FUNCTION_BLOCK Mixing
VAR_INPUT
	diEnabled : BOOL;
	iSecImp : BOOL;
END_VAR
VAR_OUTPUT
	doEnabled : BOOL;
END_VAR
VAR_IN_OUT
	MixingPhase : TPhaseMixing;
	MixerEng : TEngine;
END_VAR
VAR
	rtSecImp : R_TRIG;          // rising edge of second impulse
END_VAR

{region "Aut/Man"}
    // switching state of phase - automatic or manual control (default state is manual)
    // if both commands come at once, manual has priority (safety)
    IF MixingPhase.Cmd.ManCtrl THEN
        MixingPhase.State.ManCtrl := TRUE;
        MixingPhase.State.AutCtrl := FALSE;
    ELSIF MixingPhase.Cmd.AutCtrl THEN
        MixingPhase.State.ManCtrl := FALSE;
        MixingPhase.State.AutCtrl := TRUE;
    END_IF;

    // initialization - if neither mode is active, use manual
    IF NOT MixingPhase.State.AutCtrl AND NOT MixingPhase.State.ManCtrl THEN
        MixingPhase.State.ManCtrl := TRUE;
    END_IF;

    // commands are always reset after processing
    MixingPhase.Cmd.ManCtrl := FALSE;
    MixingPhase.Cmd.AutCtrl := FALSE;
{endregion}

{region "ManCtrl"}
    // processing manual actions - if command is processed, it is set to FALSE even if can't be processed
    // Phase commands are start, stop, pause and resume
    // Start  - start mixing (elapsed time starts from 0)
    // Stop   - stop mixing
    // Pause  - stop mixing (elapsed time is kept)
    // Resume - start mixing (continues for the remaining time)
    IF MixingPhase.State.ManCtrl THEN
        IF MixingPhase.State.Idle AND MixingPhase.Cmd.StartMan THEN
            MixingPhase.State.Running := TRUE;
            MixingPhase.State.Idle := FALSE;
            MixingPhase.State.Paused := FALSE;
            MixingPhase.State.Done := FALSE;
            MixingPhase.ElapsedTimeSec := 0;
        ELSIF MixingPhase.Cmd.StopMan THEN
            MixingPhase.State.Running := FALSE;
            MixingPhase.State.Idle := TRUE;
            MixingPhase.State.Paused := FALSE;
        ELSIF MixingPhase.State.Running AND MixingPhase.Cmd.PauseMan THEN
            MixingPhase.State.Running := FALSE;
            MixingPhase.State.Idle := FALSE;
            MixingPhase.State.Paused := TRUE;
        ELSIF MixingPhase.State.Paused AND MixingPhase.Cmd.ResumeMan THEN
            MixingPhase.State.Running := TRUE;
            MixingPhase.State.Idle := FALSE;
            MixingPhase.State.Paused := FALSE;
            MixingPhase.State.Done := FALSE;
        END_IF;
    END_IF;

    MixingPhase.Cmd.StartMan := FALSE;
    MixingPhase.Cmd.StopMan := FALSE;
    MixingPhase.Cmd.PauseMan := FALSE;
    MixingPhase.Cmd.ResumeMan := FALSE;
{endregion}

{region "AutCtrl"}
    // if phase is in automatic mode, process StartAut / StopAut (from MES)
    // commands are set to FALSE after their processing
    IF MixingPhase.State.AutCtrl THEN
        IF MixingPhase.State.Idle AND MixingPhase.Cmd.StartAut THEN
            MixingPhase.State.Running := TRUE;
            MixingPhase.State.Idle := FALSE;
            MixingPhase.State.Done := FALSE;
            MixingPhase.ElapsedTimeSec := 0;
        ELSIF MixingPhase.Cmd.StopAut THEN
            MixingPhase.State.Running := FALSE;
            MixingPhase.State.Idle := TRUE;
            MixingPhase.State.Paused := FALSE;
        END_IF;
    END_IF;

    MixingPhase.Cmd.StartAut := FALSE;
    MixingPhase.Cmd.StopAut := FALSE;
{endregion}

{region "Done"}
    // every phase should have finish condition - mixing phase - elapsed running time >= requested time
    // elapsed time is counted only while running (second impulse rising edge),
    // it is kept during pause and reset only on start
    rtSecImp(CLK := iSecImp);   // must be called every cycle, otherwise edges are lost

    IF MixingPhase.State.Running AND rtSecImp.Q THEN
        MixingPhase.ElapsedTimeSec := MixingPhase.ElapsedTimeSec + 1;
    END_IF;

    // finish condition met -> stop phase (processed next cycle) and signal Done
    IF MixingPhase.State.Running AND (MixingPhase.ElapsedTimeSec >= MixingPhase.ParamTimeSec) THEN
        MixingPhase.Cmd.StopMan := TRUE;
        MixingPhase.Cmd.StopAut := TRUE;
        MixingPhase.State.Done := TRUE;
    END_IF;

    // command reset done resets done state and then resets command
    IF MixingPhase.Cmd.ResetDone THEN
        MixingPhase.State.Done := FALSE;
        MixingPhase.Cmd.ResetDone := FALSE;
    END_IF;
{endregion}

{region "States"}
    // Command mixer in cases of states
    // Running - mixer runs
    // Idle    - mixer stopped
    // Paused  - mixer stopped
    IF MixingPhase.State.Running THEN
        MixerEng.Cmd.Req2RunAutCtrl := TRUE;
    ELSE
        MixerEng.Cmd.Req2RunAutCtrl := FALSE;
    END_IF;
{endregion}

// default state of phase - if not any state sets state to idle
IF NOT MixingPhase.State.Idle AND NOT MixingPhase.State.Paused AND NOT MixingPhase.State.Running THEN
    MixingPhase.State.Idle := 1;
END_IF;

// write binary states into int value for visualization
IF MixingPhase.State.Idle THEN
    MixingPhase.State.Stateint := Global.PhIdle;
ELSIF MixingPhase.State.Running THEN
    MixingPhase.State.Stateint := Global.PhRunning;
ELSE
    MixingPhase.State.Stateint := Global.PhPause;
END_IF;

doEnabled := diEnabled;

END_FUNCTION_BLOCK

(* stored: Version 1.1.0.1, ProductVersion 3.1.4026.21
   POU Mixing: Id {c7d77201-326e-43f5-84be-5e5d3f37b70d}, SpecialFunc None *)
